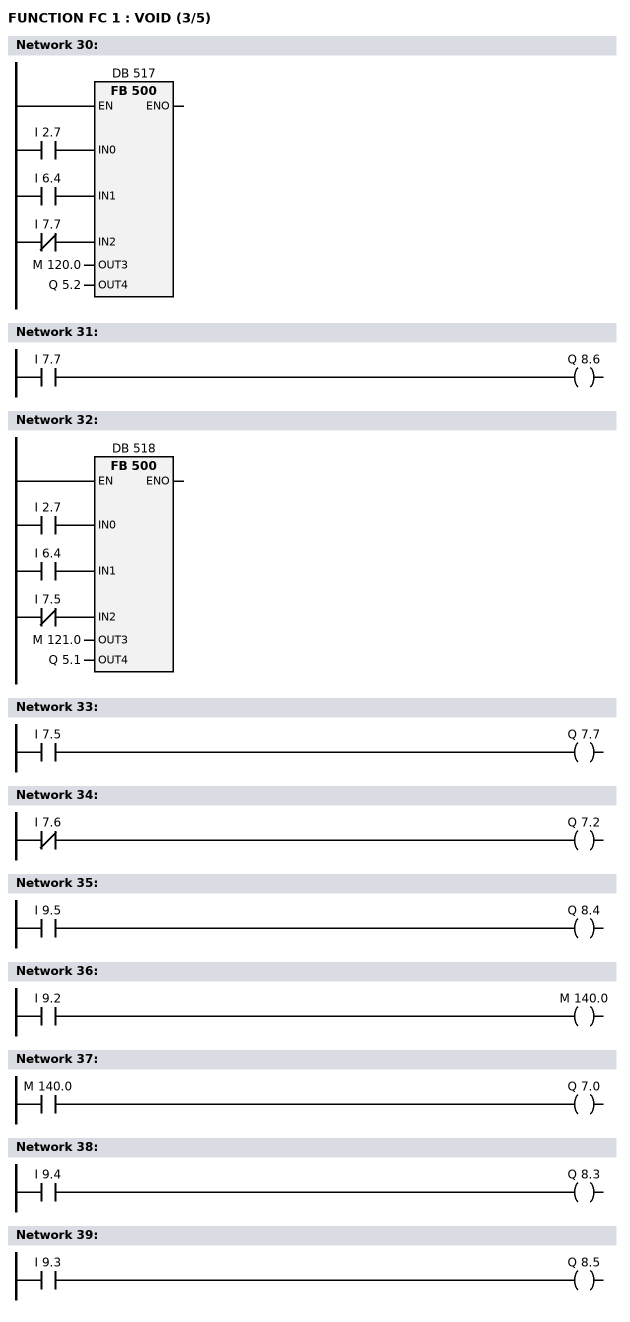

      A     I      2.7;
      =     L      0.0;
      BLD   103;
      A     I      6.4;
      =     L      0.1;
      BLD   103;
      AN    I      7.7;
      =     L      0.2;
      BLD   103;
      CALL FB   500 , DB   517 (
           IN0                      := L      0.0,
           IN1                      := L      0.1,
           IN2                      := L      0.2,
           OUT3                     := M    120.0,
           OUT4                     := Q      5.2);
      NOP   0;
NETWORK
TITLE =

      A     I      7.7;
      =     Q      8.6;
NETWORK
TITLE =

      A     I      2.7;
      =     L      0.0;
      BLD   103;
      A     I      6.4;
      =     L      0.1;
      BLD   103;
      AN    I      7.5;
      =     L      0.2;
      BLD   103;
      CALL FB   500 , DB   518 (
           IN0                      := L      0.0,
           IN1                      := L      0.1,
           IN2                      := L      0.2,
           OUT3                     := M    121.0,
           OUT4                     := Q      5.1);
      NOP   0;
NETWORK
TITLE =

      A     I      7.5;
      =     Q      7.7;
NETWORK
TITLE =

      AN    I      7.6;
      =     Q      7.2;
NETWORK
TITLE =

      A     I      9.5;
      =     Q      8.4;
NETWORK
TITLE =

      A     I      9.2;
      =     M    140.0;
NETWORK
TITLE =

      A     M    140.0;
      =     Q      7.0;
NETWORK
TITLE =

      A     I      9.4;
      =     Q      8.3;
NETWORK
TITLE =

      A     I      9.3;
      =     Q      8.5;
NETWORK
TITLE =
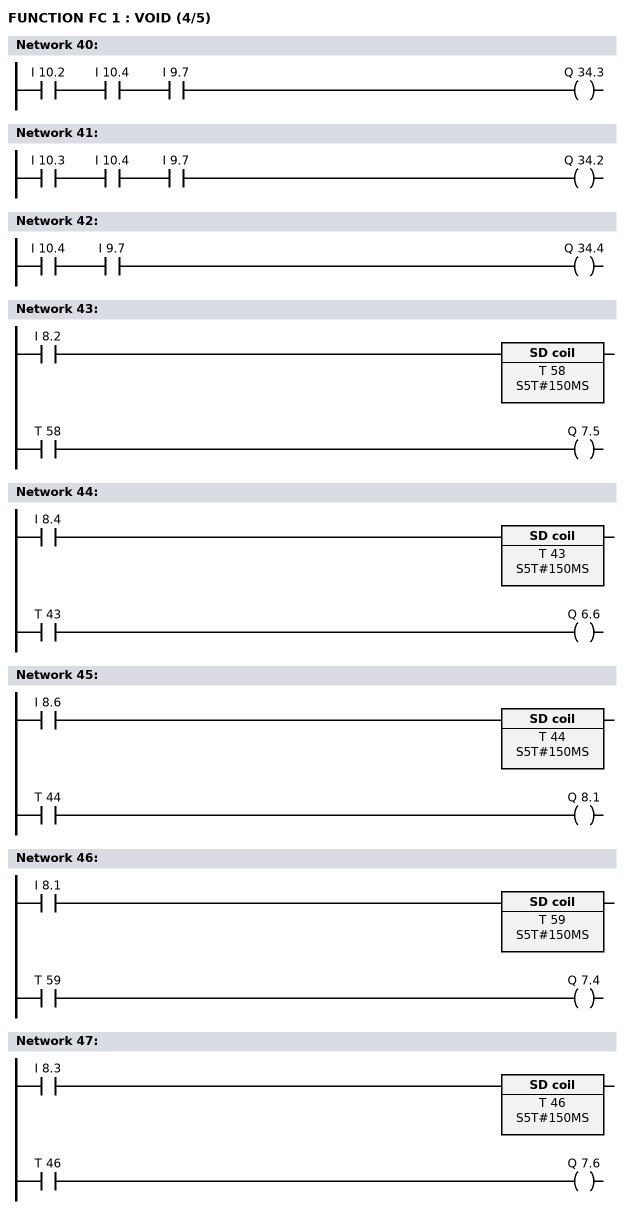

      A     I     10.2;
      A     I     10.4;
      A     I      9.7;
      =     Q     34.3;
NETWORK
TITLE =

      A     I     10.3;
      A     I     10.4;
      A     I      9.7;
      =     Q     34.2;
NETWORK
TITLE =

      A     I     10.4;
      A     I      9.7;
      =     Q     34.4;
NETWORK
TITLE =

      A     I      8.2;
      L     S5T#150MS;
      SD    T     58;
      NOP   0;
      NOP   0;
      NOP   0;
      A     T     58;
      =     Q      7.5;
NETWORK
TITLE =

      A     I      8.4;
      L     S5T#150MS;
      SD    T     43;
      NOP   0;
      NOP   0;
      NOP   0;
      A     T     43;
      =     Q      6.6;
NETWORK
TITLE =

      A     I      8.6;
      L     S5T#150MS;
      SD    T     44;
      NOP   0;
      NOP   0;
      NOP   0;
      A     T     44;
      =     Q      8.1;
NETWORK
TITLE =

      A     I      8.1;
      L     S5T#150MS;
      SD    T     59;
      NOP   0;
      NOP   0;
      NOP   0;
      A     T     59;
      =     Q      7.4;
NETWORK
TITLE =

      A     I      8.3;
      L     S5T#150MS;
      SD    T     46;
      NOP   0;
      NOP   0;
      NOP   0;
      A     T     46;
      =     Q      7.6;
NETWORK
TITLE =
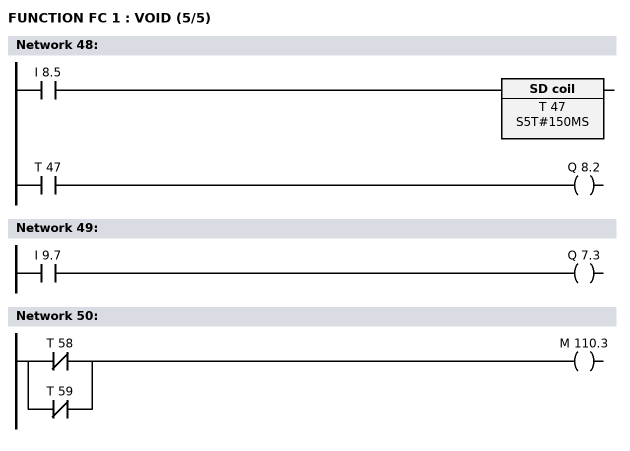

      A     I      8.5;
      L     S5T#150MS;
      SD    T     47;
      NOP   0;
      NOP   0;
      NOP   0;
      A     T     47;
      =     Q      8.2;
NETWORK
TITLE =

      A     I      9.7;
      =     Q      7.3;
NETWORK
TITLE =

      ON    T     58;
      ON    T     59;
      =     M    110.3;
END_FUNCTION

FUNCTION FC 2 : VOID
VERSION : 0.1

BEGIN
NETWORK
TITLE =
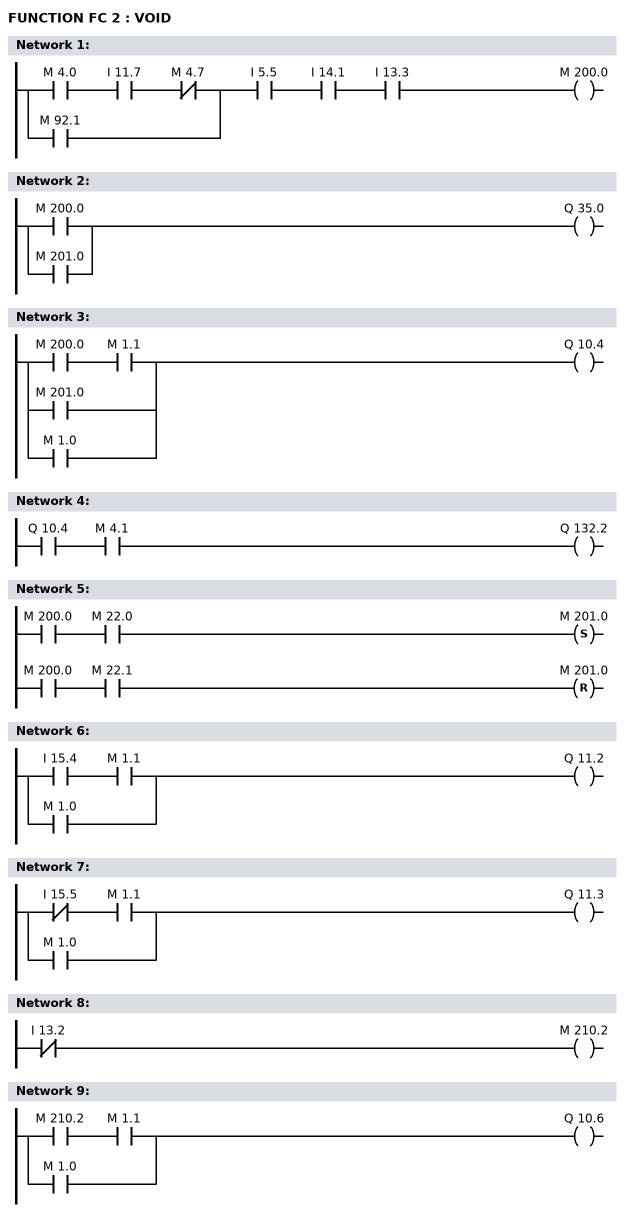

      A(    ;
      A     M      4.0;
      A     I     11.7;
      AN    M      4.7;
      O     M     92.1;
      )     ;
      A     I      5.5;
      A     I     14.1;
      A     I     13.3;
      =     M    200.0;
NETWORK
TITLE =

      O     M    200.0;
      O     M    201.0;
      =     Q     35.0;
NETWORK
TITLE =

      A     M    200.0;
      A     M      1.1;
      O     M    201.0;
      O     M      1.0;
      =     Q     10.4;
NETWORK
TITLE =

      A     Q     10.4;
      A     M      4.1;
      =     Q    132.2;
NETWORK
TITLE =

      A     M    200.0;
      A     M     22.0;
      S     M    201.0;
      A     M    200.0;
      A     M     22.1;
      R     M    201.0;
      NOP   0;
NETWORK
TITLE =

      A     I     15.4;
      A     M      1.1;
      O     M      1.0;
      =     Q     11.2;
NETWORK
TITLE =

      AN    I     15.5;
      A     M      1.1;
      O     M      1.0;
      =     Q     11.3;
NETWORK
TITLE =

      AN    I     13.2;
      =     M    210.2;
NETWORK
TITLE =

      A     M    210.2;
      A     M      1.1;
      O     M      1.0;
      =     Q     10.6;
NETWORK
TITLE =

      O(    ;
      A     I     12.3;
      L     S5T#150MS;
      SD    T     70;
      NOP   0;
      NOP   0;
      NOP   0;
      A     T     70;
      )     ;
      O     M      1.0;
      =     Q     10.3;
NETWORK
TITLE =
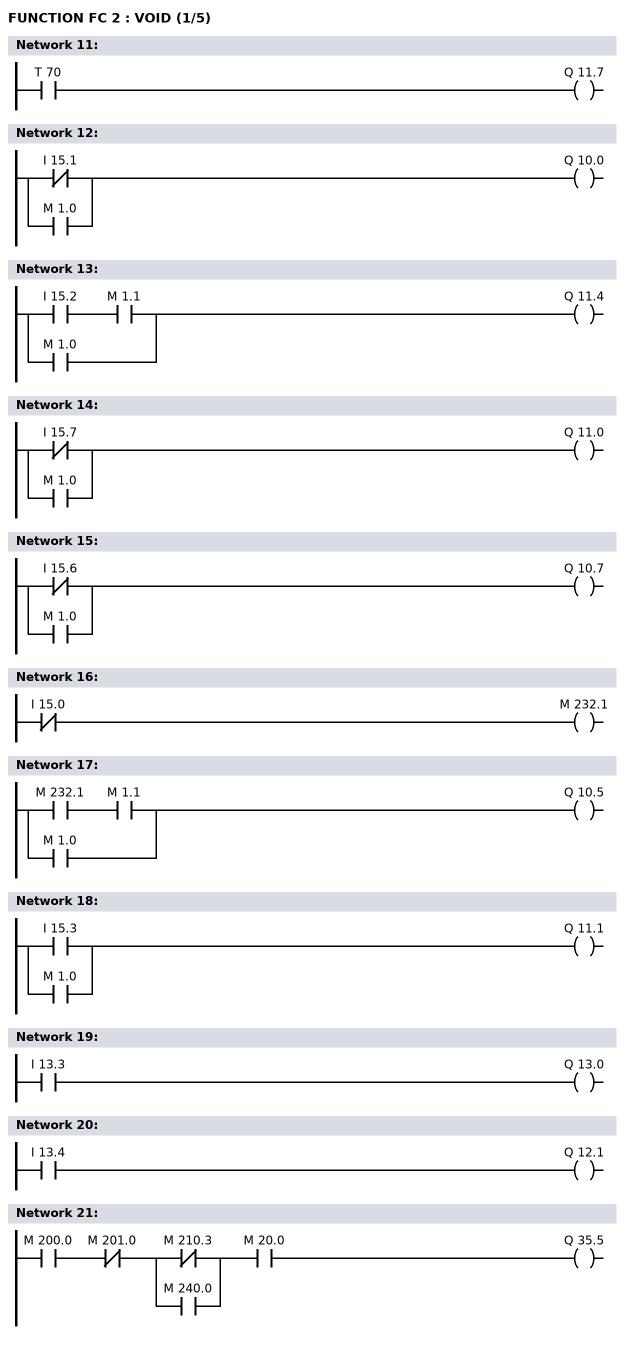

      A     T     70;
      =     Q     11.7;
NETWORK
TITLE =

      ON    I     15.1;
      O     M      1.0;
      =     Q     10.0;
NETWORK
TITLE =

      A     I     15.2;
      A     M      1.1;
      O     M      1.0;
      =     Q     11.4;
NETWORK
TITLE =

      ON    I     15.7;
      O     M      1.0;
      =     Q     11.0;
NETWORK
TITLE =

      ON    I     15.6;
      O     M      1.0;
      =     Q     10.7;
NETWORK
TITLE =

      AN    I     15.0;
      =     M    232.1;
NETWORK
TITLE =

      A     M    232.1;
      A     M      1.1;
      O     M      1.0;
      =     Q     10.5;
NETWORK
TITLE =

      O     I     15.3;
      O     M      1.0;
      =     Q     11.1;
NETWORK
TITLE =

      A     I     13.3;
      =     Q     13.0;
NETWORK
TITLE =

      A     I     13.4;
      =     Q     12.1;
NETWORK
TITLE =

      A     M    200.0;
      AN    M    201.0;
      A(    ;
      ON    M    210.3;
      O     M    240.0;
      )     ;
      A     M     20.0;
      =     Q     35.5;
NETWORK
TITLE =
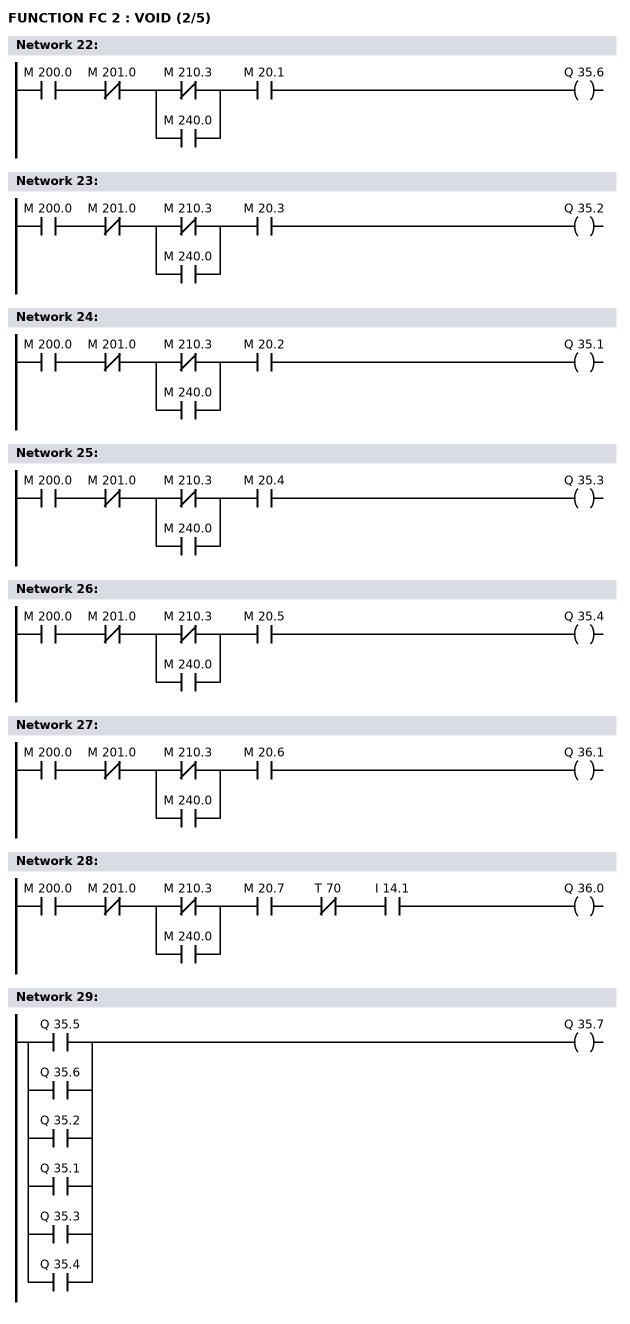

      A     M    200.0;
      AN    M    201.0;
      A(    ;
      ON    M    210.3;
      O     M    240.0;
      )     ;
      A     M     20.1;
      =     Q     35.6;
NETWORK
TITLE =

      A     M    200.0;
      AN    M    201.0;
      A(    ;
      ON    M    210.3;
      O     M    240.0;
      )     ;
      A     M     20.3;
      =     Q     35.2;
NETWORK
TITLE =

      A     M    200.0;
      AN    M    201.0;
      A(    ;
      ON    M    210.3;
      O     M    240.0;
      )     ;
      A     M     20.2;
      =     Q     35.1;
NETWORK
TITLE =

      A     M    200.0;
      AN    M    201.0;
      A(    ;
      ON    M    210.3;
      O     M    240.0;
      )     ;
      A     M     20.4;
      =     Q     35.3;
NETWORK
TITLE =

      A     M    200.0;
      AN    M    201.0;
      A(    ;
      ON    M    210.3;
      O     M    240.0;
      )     ;
      A     M     20.5;
      =     Q     35.4;
NETWORK
TITLE =

      A     M    200.0;
      AN    M    201.0;
      A(    ;
      ON    M    210.3;
      O     M    240.0;
      )     ;
      A     M     20.6;
      =     Q     36.1;
NETWORK
TITLE =

      A     M    200.0;
      AN    M    201.0;
      A(    ;
      ON    M    210.3;
      O     M    240.0;
      )     ;
      A     M     20.7;
      AN    T     70;
      A     I     14.1;
      =     Q     36.0;
NETWORK
TITLE =

      O     Q     35.5;
      O     Q     35.6;
      O     Q     35.2;
      O     Q     35.1;
      O     Q     35.3;
      O     Q     35.4;
      =     Q     35.7;
NETWORK
TITLE =
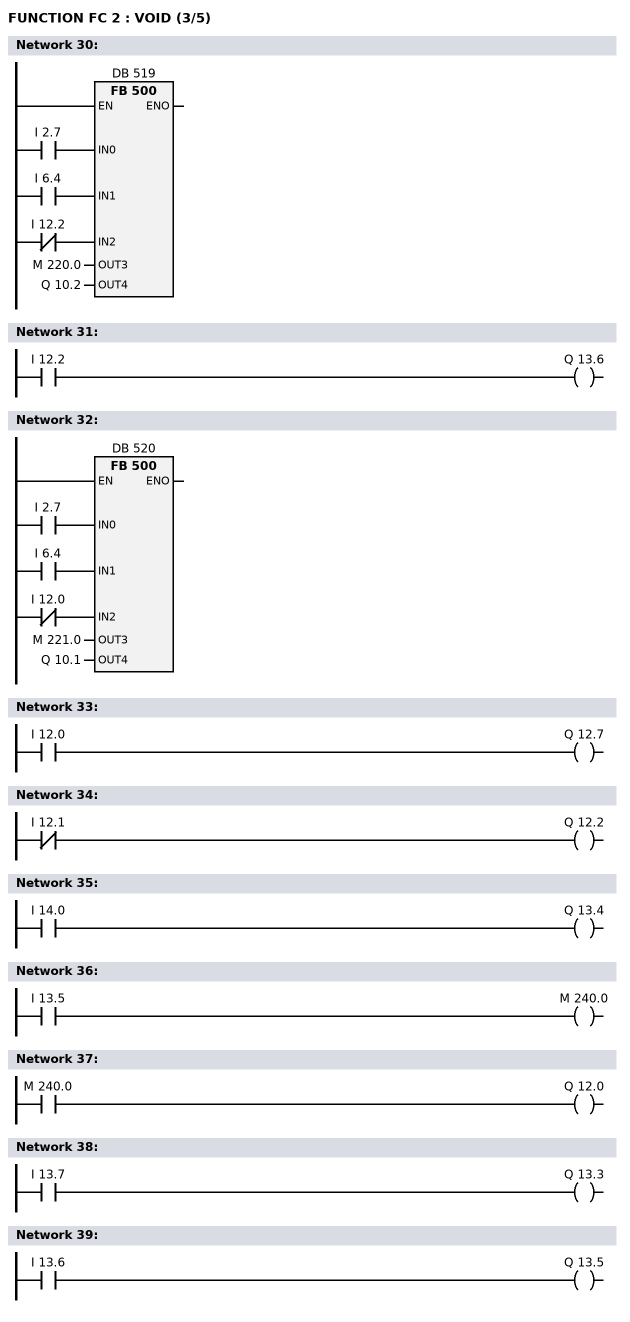

      A     I      2.7;
      =     L      0.0;
      BLD   103;
      A     I      6.4;
      =     L      0.1;
      BLD   103;
      AN    I     12.2;
      =     L      0.2;
      BLD   103;
      CALL FB   500 , DB   519 (
           IN0                      := L      0.0,
           IN1                      := L      0.1,
           IN2                      := L      0.2,
           OUT3                     := M    220.0,
           OUT4                     := Q     10.2);
      NOP   0;
NETWORK
TITLE =

      A     I     12.2;
      =     Q     13.6;
NETWORK
TITLE =

      A     I      2.7;
      =     L      0.0;
      BLD   103;
      A     I      6.4;
      =     L      0.1;
      BLD   103;
      AN    I     12.0;
      =     L      0.2;
      BLD   103;
      CALL FB   500 , DB   520 (
           IN0                      := L      0.0,
           IN1                      := L      0.1,
           IN2                      := L      0.2,
           OUT3                     := M    221.0,
           OUT4                     := Q     10.1);
      NOP   0;
NETWORK
TITLE =

      A     I     12.0;
      =     Q     12.7;
NETWORK
TITLE =

      AN    I     12.1;
      =     Q     12.2;
NETWORK
TITLE =

      A     I     14.0;
      =     Q     13.4;
NETWORK
TITLE =

      A     I     13.5;
      =     M    240.0;
NETWORK
TITLE =

      A     M    240.0;
      =     Q     12.0;
NETWORK
TITLE =

      A     I     13.7;
      =     Q     13.3;
NETWORK
TITLE =

      A     I     13.6;
      =     Q     13.5;
NETWORK
TITLE =
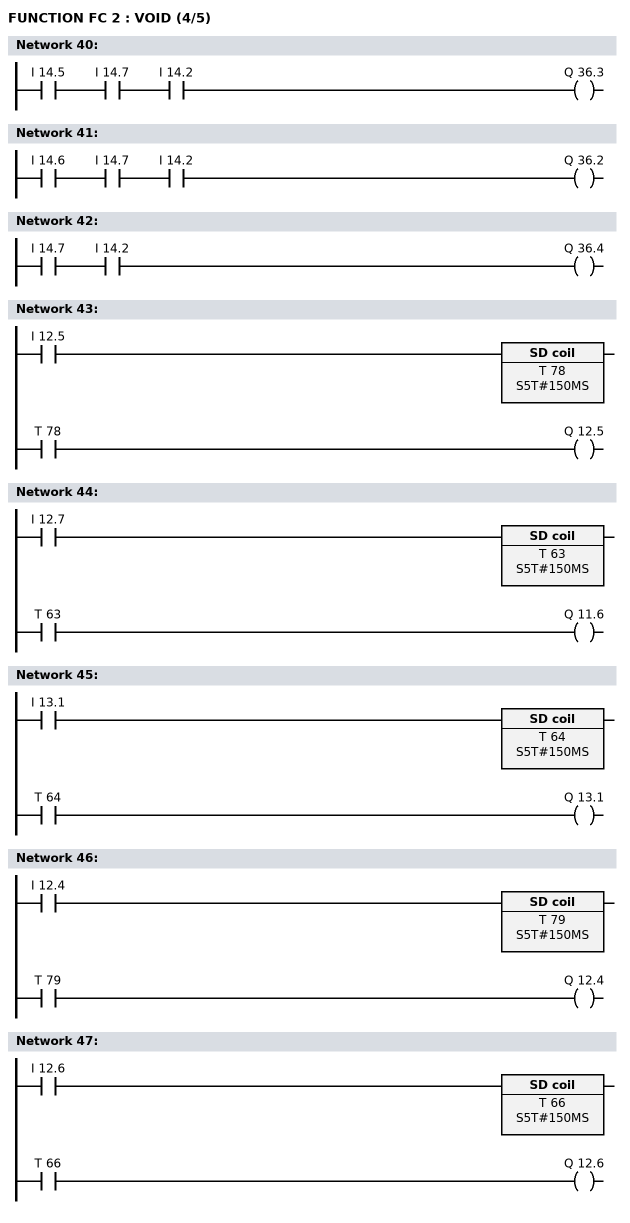

      A     I     14.5;
      A     I     14.7;
      A     I     14.2;
      =     Q     36.3;
NETWORK
TITLE =

      A     I     14.6;
      A     I     14.7;
      A     I     14.2;
      =     Q     36.2;
NETWORK
TITLE =

      A     I     14.7;
      A     I     14.2;
      =     Q     36.4;
NETWORK
TITLE =

      A     I     12.5;
      L     S5T#150MS;
      SD    T     78;
      NOP   0;
      NOP   0;
      NOP   0;
      A     T     78;
      =     Q     12.5;
NETWORK
TITLE =

      A     I     12.7;
      L     S5T#150MS;
      SD    T     63;
      NOP   0;
      NOP   0;
      NOP   0;
      A     T     63;
      =     Q     11.6;
NETWORK
TITLE =

      A     I     13.1;
      L     S5T#150MS;
      SD    T     64;
      NOP   0;
      NOP   0;
      NOP   0;
      A     T     64;
      =     Q     13.1;
NETWORK
TITLE =

      A     I     12.4;
      L     S5T#150MS;
      SD    T     79;
      NOP   0;
      NOP   0;
      NOP   0;
      A     T     79;
      =     Q     12.4;
NETWORK
TITLE =

      A     I     12.6;
      L     S5T#150MS;
      SD    T     66;
      NOP   0;
      NOP   0;
      NOP   0;
      A     T     66;
      =     Q     12.6;
NETWORK
TITLE =
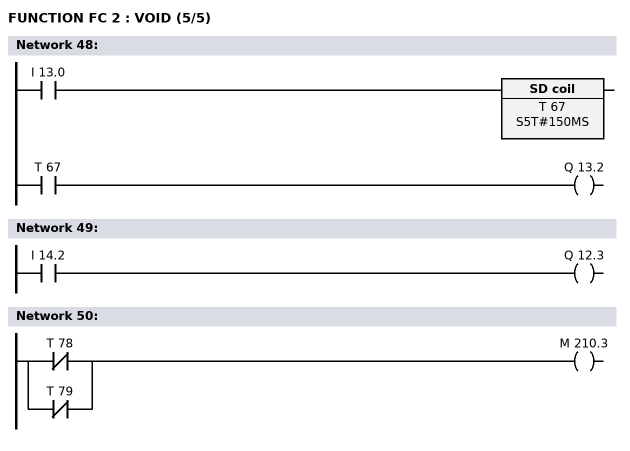

      A     I     13.0;
      L     S5T#150MS;
      SD    T     67;
      NOP   0;
      NOP   0;
      NOP   0;
      A     T     67;
      =     Q     13.2;
NETWORK
TITLE =

      A     I     14.2;
      =     Q     12.3;
NETWORK
TITLE =

      ON    T     78;
      ON    T     79;
      =     M    210.3;
END_FUNCTION

FUNCTION FC 3 : VOID
VERSION : 0.1

BEGIN
NETWORK
TITLE =
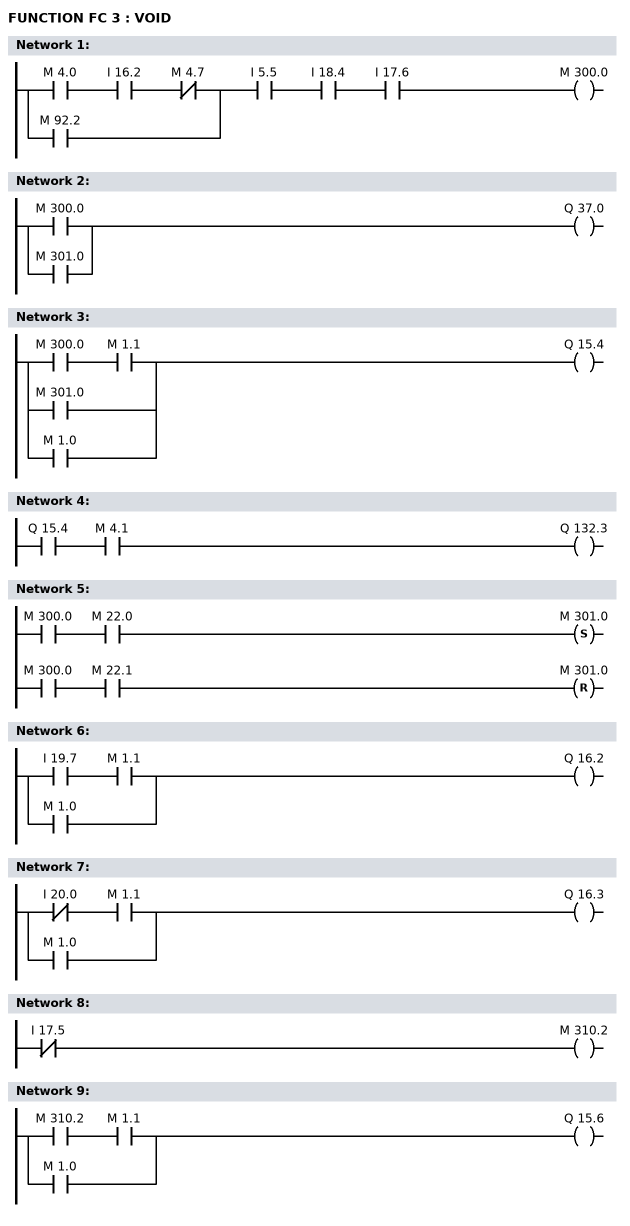

      A(    ;
      A     M      4.0;
      A     I     16.2;
      AN    M      4.7;
      O     M     92.2;
      )     ;
      A     I      5.5;
      A     I     18.4;
      A     I     17.6;
      =     M    300.0;
NETWORK
TITLE =

      O     M    300.0;
      O     M    301.0;
      =     Q     37.0;
NETWORK
TITLE =

      A     M    300.0;
      A     M      1.1;
      O     M    301.0;
      O     M      1.0;
      =     Q     15.4;
NETWORK
TITLE =

      A     Q     15.4;
      A     M      4.1;
      =     Q    132.3;
NETWORK
TITLE =

      A     M    300.0;
      A     M     22.0;
      S     M    301.0;
      A     M    300.0;
      A     M     22.1;
      R     M    301.0;
      NOP   0;
NETWORK
TITLE =

      A     I     19.7;
      A     M      1.1;
      O     M      1.0;
      =     Q     16.2;
NETWORK
TITLE =

      AN    I     20.0;
      A     M      1.1;
      O     M      1.0;
      =     Q     16.3;
NETWORK
TITLE =

      AN    I     17.5;
      =     M    310.2;
NETWORK
TITLE =

      A     M    310.2;
      A     M      1.1;
      O     M      1.0;
      =     Q     15.6;
NETWORK
TITLE =

      O(    ;
      A     I     16.6;
      L     S5T#150MS;
      SD    T     90;
      NOP   0;
      NOP   0;
      NOP   0;
      A     T     90;
      )     ;
      O     M      1.0;
      =     Q     15.3;
NETWORK
TITLE =
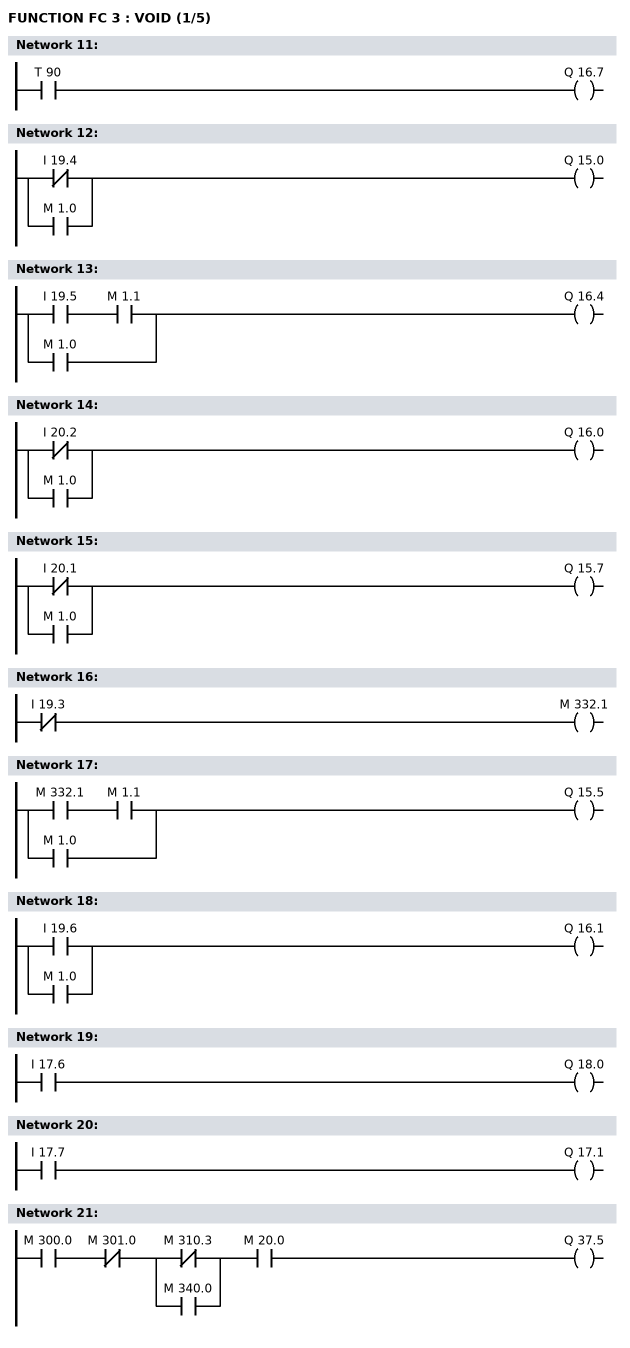

      A     T     90;
      =     Q     16.7;
NETWORK
TITLE =

      ON    I     19.4;
      O     M      1.0;
      =     Q     15.0;
NETWORK
TITLE =

      A     I     19.5;
      A     M      1.1;
      O     M      1.0;
      =     Q     16.4;
NETWORK
TITLE =

      ON    I     20.2;
      O     M      1.0;
      =     Q     16.0;
NETWORK
TITLE =

      ON    I     20.1;
      O     M      1.0;
      =     Q     15.7;
NETWORK
TITLE =

      AN    I     19.3;
      =     M    332.1;
NETWORK
TITLE =

      A     M    332.1;
      A     M      1.1;
      O     M      1.0;
      =     Q     15.5;
NETWORK
TITLE =

      O     I     19.6;
      O     M      1.0;
      =     Q     16.1;
NETWORK
TITLE =

      A     I     17.6;
      =     Q     18.0;
NETWORK
TITLE =

      A     I     17.7;
      =     Q     17.1;
NETWORK
TITLE =

      A     M    300.0;
      AN    M    301.0;
      A(    ;
      ON    M    310.3;
      O     M    340.0;
      )     ;
      A     M     20.0;
      =     Q     37.5;
NETWORK
TITLE =
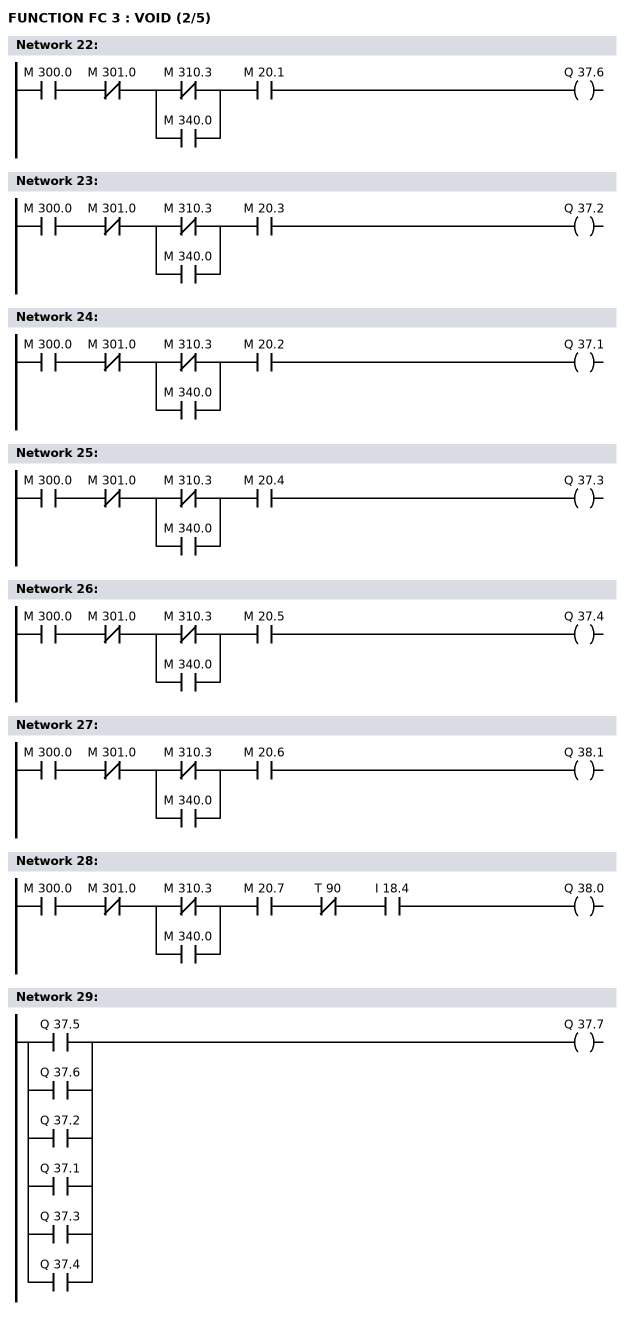

      A     M    300.0;
      AN    M    301.0;
      A(    ;
      ON    M    310.3;
      O     M    340.0;
      )     ;
      A     M     20.1;
      =     Q     37.6;
NETWORK
TITLE =

      A     M    300.0;
      AN    M    301.0;
      A(    ;
      ON    M    310.3;
      O     M    340.0;
      )     ;
      A     M     20.3;
      =     Q     37.2;
NETWORK
TITLE =

      A     M    300.0;
      AN    M    301.0;
      A(    ;
      ON    M    310.3;
      O     M    340.0;
      )     ;
      A     M     20.2;
      =     Q     37.1;
NETWORK
TITLE =

      A     M    300.0;
      AN    M    301.0;
      A(    ;
      ON    M    310.3;
      O     M    340.0;
      )     ;
      A     M     20.4;
      =     Q     37.3;
NETWORK
TITLE =

      A     M    300.0;
      AN    M    301.0;
      A(    ;
      ON    M    310.3;
      O     M    340.0;
      )     ;
      A     M     20.5;
      =     Q     37.4;
NETWORK
TITLE =

      A     M    300.0;
      AN    M    301.0;
      A(    ;
      ON    M    310.3;
      O     M    340.0;
      )     ;
      A     M     20.6;
      =     Q     38.1;
NETWORK
TITLE =

      A     M    300.0;
      AN    M    301.0;
      A(    ;
      ON    M    310.3;
      O     M    340.0;
      )     ;
      A     M     20.7;
      AN    T     90;
      A     I     18.4;
      =     Q     38.0;
NETWORK
TITLE =

      O     Q     37.5;
      O     Q     37.6;
      O     Q     37.2;
      O     Q     37.1;
      O     Q     37.3;
      O     Q     37.4;
      =     Q     37.7;
NETWORK
TITLE =
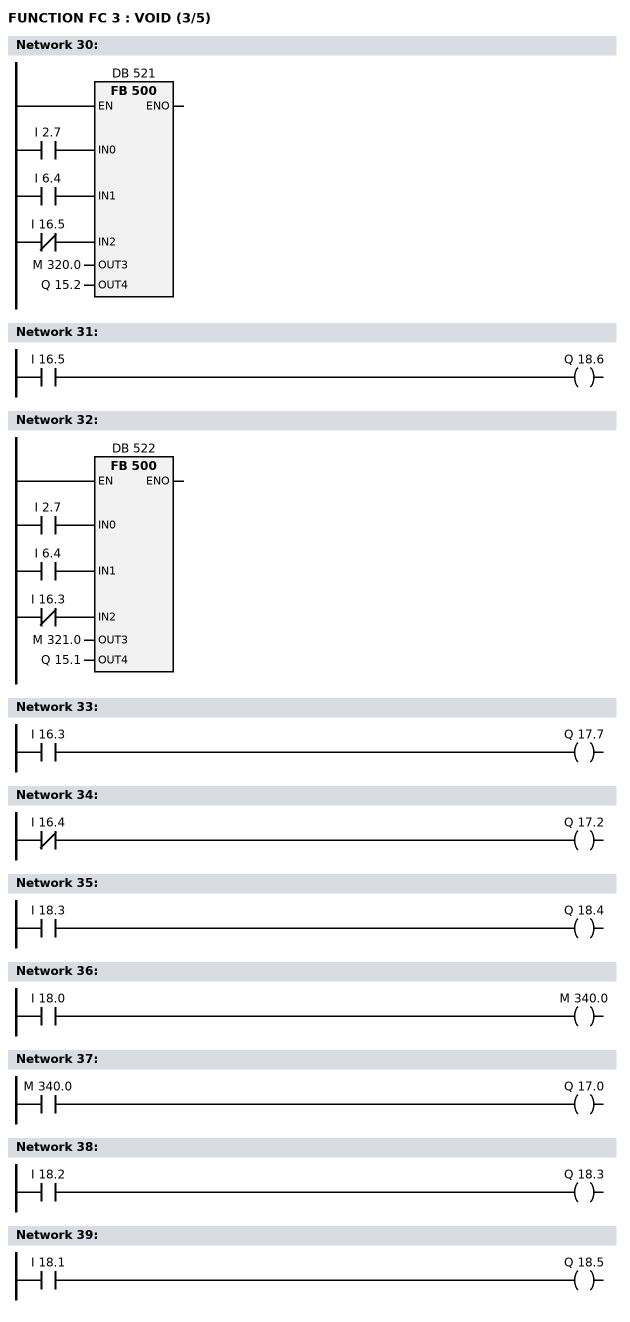

      A     I      2.7;
      =     L      0.0;
      BLD   103;
      A     I      6.4;
      =     L      0.1;
      BLD   103;
      AN    I     16.5;
      =     L      0.2;
      BLD   103;
      CALL FB   500 , DB   521 (
           IN0                      := L      0.0,
           IN1                      := L      0.1,
           IN2                      := L      0.2,
           OUT3                     := M    320.0,
           OUT4                     := Q     15.2);
      NOP   0;
NETWORK
TITLE =

      A     I     16.5;
      =     Q     18.6;
NETWORK
TITLE =

      A     I      2.7;
      =     L      0.0;
      BLD   103;
      A     I      6.4;
      =     L      0.1;
      BLD   103;
      AN    I     16.3;
      =     L      0.2;
      BLD   103;
      CALL FB   500 , DB   522 (
           IN0                      := L      0.0,
           IN1                      := L      0.1,
           IN2                      := L      0.2,
           OUT3                     := M    321.0,
           OUT4                     := Q     15.1);
      NOP   0;
NETWORK
TITLE =

      A     I     16.3;
      =     Q     17.7;
NETWORK
TITLE =

      AN    I     16.4;
      =     Q     17.2;
NETWORK
TITLE =

      A     I     18.3;
      =     Q     18.4;
NETWORK
TITLE =

      A     I     18.0;
      =     M    340.0;
NETWORK
TITLE =

      A     M    340.0;
      =     Q     17.0;
NETWORK
TITLE =

      A     I     18.2;
      =     Q     18.3;
NETWORK
TITLE =

      A     I     18.1;
      =     Q     18.5;
NETWORK
TITLE =
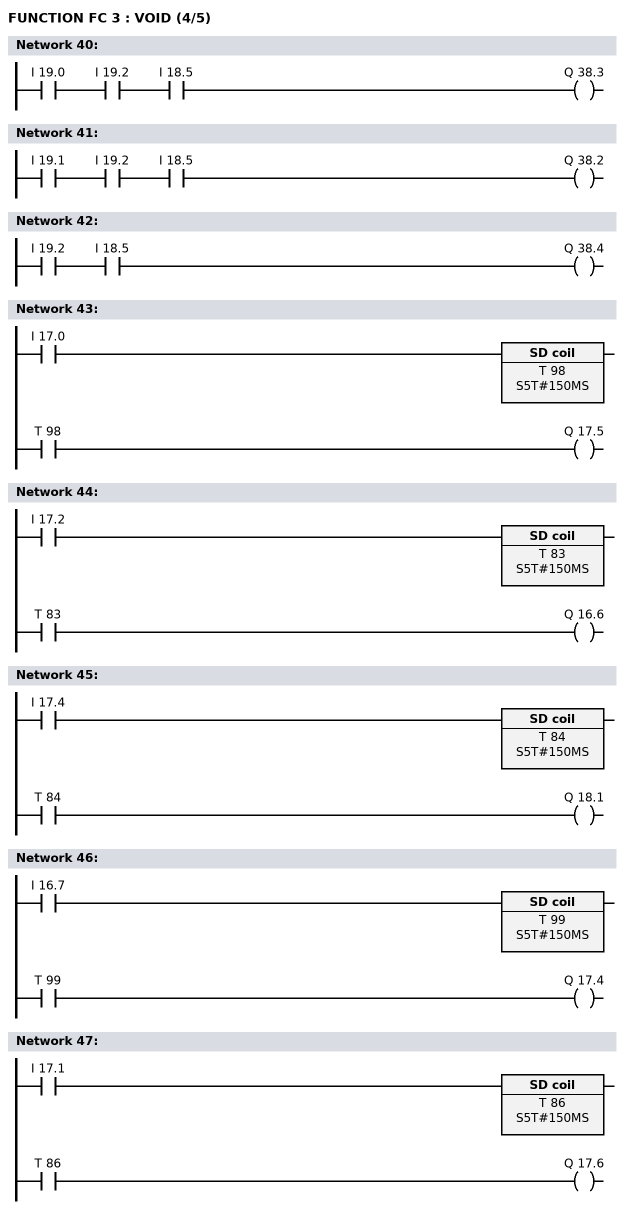

      A     I     19.0;
      A     I     19.2;
      A     I     18.5;
      =     Q     38.3;
NETWORK
TITLE =

      A     I     19.1;
      A     I     19.2;
      A     I     18.5;
      =     Q     38.2;
NETWORK
TITLE =

      A     I     19.2;
      A     I     18.5;
      =     Q     38.4;
NETWORK
TITLE =

      A     I     17.0;
      L     S5T#150MS;
      SD    T     98;
      NOP   0;
      NOP   0;
      NOP   0;
      A     T     98;
      =     Q     17.5;
NETWORK
TITLE =

      A     I     17.2;
      L     S5T#150MS;
      SD    T     83;
      NOP   0;
      NOP   0;
      NOP   0;
      A     T     83;
      =     Q     16.6;
NETWORK
TITLE =

      A     I     17.4;
      L     S5T#150MS;
      SD    T     84;
      NOP   0;
      NOP   0;
      NOP   0;
      A     T     84;
      =     Q     18.1;
NETWORK
TITLE =

      A     I     16.7;
      L     S5T#150MS;
      SD    T     99;
      NOP   0;
      NOP   0;
      NOP   0;
      A     T     99;
      =     Q     17.4;
NETWORK
TITLE =

      A     I     17.1;
      L     S5T#150MS;
      SD    T     86;
      NOP   0;
      NOP   0;
      NOP   0;
      A     T     86;
      =     Q     17.6;
NETWORK
TITLE =
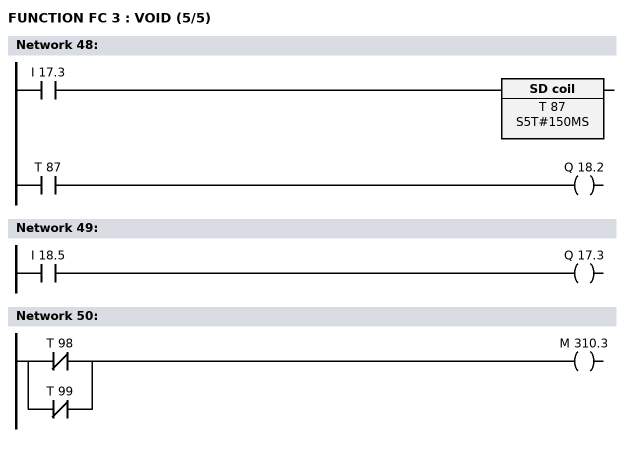

      A     I     17.3;
      L     S5T#150MS;
      SD    T     87;
      NOP   0;
      NOP   0;
      NOP   0;
      A     T     87;
      =     Q     18.2;
NETWORK
TITLE =

      A     I     18.5;
      =     Q     17.3;
NETWORK
TITLE =

      ON    T     98;
      ON    T     99;
      =     M    310.3;
END_FUNCTION

FUNCTION FC 4 : VOID
VERSION : 0.1

BEGIN
NETWORK
TITLE =
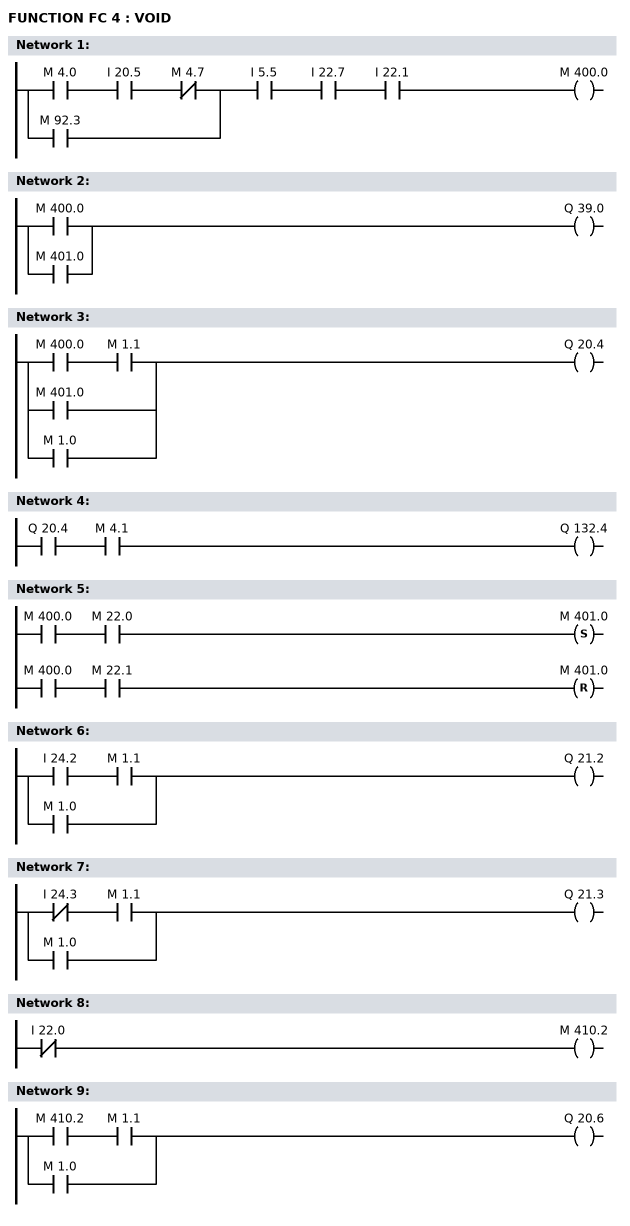

      A(    ;
      A     M      4.0;
      A     I     20.5;
      AN    M      4.7;
      O     M     92.3;
      )     ;
      A     I      5.5;
      A     I     22.7;
      A     I     22.1;
      =     M    400.0;
NETWORK
TITLE =

      O     M    400.0;
      O     M    401.0;
      =     Q     39.0;
NETWORK
TITLE =

      A     M    400.0;
      A     M      1.1;
      O     M    401.0;
      O     M      1.0;
      =     Q     20.4;
NETWORK
TITLE =

      A     Q     20.4;
      A     M      4.1;
      =     Q    132.4;
NETWORK
TITLE =

      A     M    400.0;
      A     M     22.0;
      S     M    401.0;
      A     M    400.0;
      A     M     22.1;
      R     M    401.0;
      NOP   0;
NETWORK
TITLE =

      A     I     24.2;
      A     M      1.1;
      O     M      1.0;
      =     Q     21.2;
NETWORK
TITLE =

      AN    I     24.3;
      A     M      1.1;
      O     M      1.0;
      =     Q     21.3;
NETWORK
TITLE =

      AN    I     22.0;
      =     M    410.2;
NETWORK
TITLE =

      A     M    410.2;
      A     M      1.1;
      O     M      1.0;
      =     Q     20.6;
NETWORK
TITLE =

      O(    ;
      A     I     21.1;
      L     S5T#150MS;
      SD    T    110;
      NOP   0;
      NOP   0;
      NOP   0;
      A     T    110;
      )     ;
      O     M      1.0;
      =     Q     20.3;
NETWORK
TITLE =
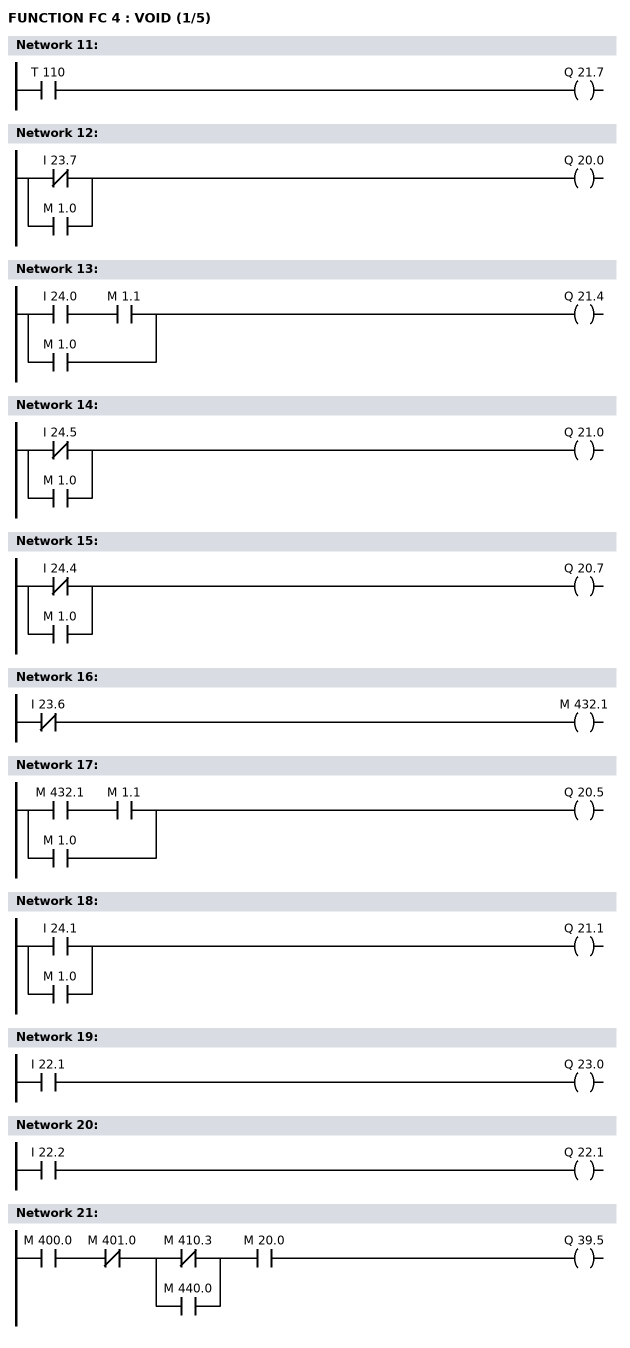

      A     T    110;
      =     Q     21.7;
NETWORK
TITLE =

      ON    I     23.7;
      O     M      1.0;
      =     Q     20.0;
NETWORK
TITLE =

      A     I     24.0;
      A     M      1.1;
      O     M      1.0;
      =     Q     21.4;
NETWORK
TITLE =

      ON    I     24.5;
      O     M      1.0;
      =     Q     21.0;
NETWORK
TITLE =

      ON    I     24.4;
      O     M      1.0;
      =     Q     20.7;
NETWORK
TITLE =

      AN    I     23.6;
      =     M    432.1;
NETWORK
TITLE =

      A     M    432.1;
      A     M      1.1;
      O     M      1.0;
      =     Q     20.5;
NETWORK
TITLE =

      O     I     24.1;
      O     M      1.0;
      =     Q     21.1;
NETWORK
TITLE =

      A     I     22.1;
      =     Q     23.0;
NETWORK
TITLE =

      A     I     22.2;
      =     Q     22.1;
NETWORK
TITLE =

      A     M    400.0;
      AN    M    401.0;
      A(    ;
      ON    M    410.3;
      O     M    440.0;
      )     ;
      A     M     20.0;
      =     Q     39.5;
NETWORK
TITLE =
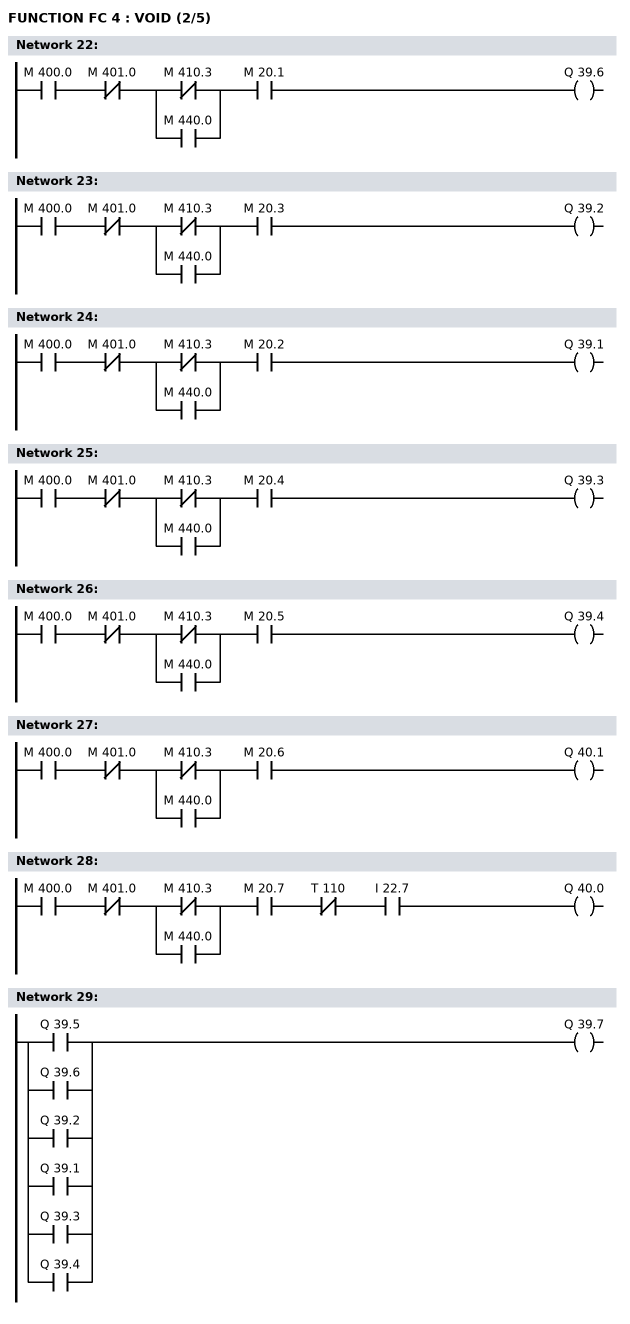

      A     M    400.0;
      AN    M    401.0;
      A(    ;
      ON    M    410.3;
      O     M    440.0;
      )     ;
      A     M     20.1;
      =     Q     39.6;
NETWORK
TITLE =

      A     M    400.0;
      AN    M    401.0;
      A(    ;
      ON    M    410.3;
      O     M    440.0;
      )     ;
      A     M     20.3;
      =     Q     39.2;
NETWORK
TITLE =

      A     M    400.0;
      AN    M    401.0;
      A(    ;
      ON    M    410.3;
      O     M    440.0;
      )     ;
      A     M     20.2;
      =     Q     39.1;
NETWORK
TITLE =

      A     M    400.0;
      AN    M    401.0;
      A(    ;
      ON    M    410.3;
      O     M    440.0;
      )     ;
      A     M     20.4;
      =     Q     39.3;
NETWORK
TITLE =

      A     M    400.0;
      AN    M    401.0;
      A(    ;
      ON    M    410.3;
      O     M    440.0;
      )     ;
      A     M     20.5;
      =     Q     39.4;
NETWORK
TITLE =

      A     M    400.0;
      AN    M    401.0;
      A(    ;
      ON    M    410.3;
      O     M    440.0;
      )     ;
      A     M     20.6;
      =     Q     40.1;
NETWORK
TITLE =

      A     M    400.0;
      AN    M    401.0;
      A(    ;
      ON    M    410.3;
      O     M    440.0;
      )     ;
      A     M     20.7;
      AN    T    110;
      A     I     22.7;
      =     Q     40.0;
NETWORK
TITLE =

      O     Q     39.5;
      O     Q     39.6;
      O     Q     39.2;
      O     Q     39.1;
      O     Q     39.3;
      O     Q     39.4;
      =     Q     39.7;
NETWORK
TITLE =
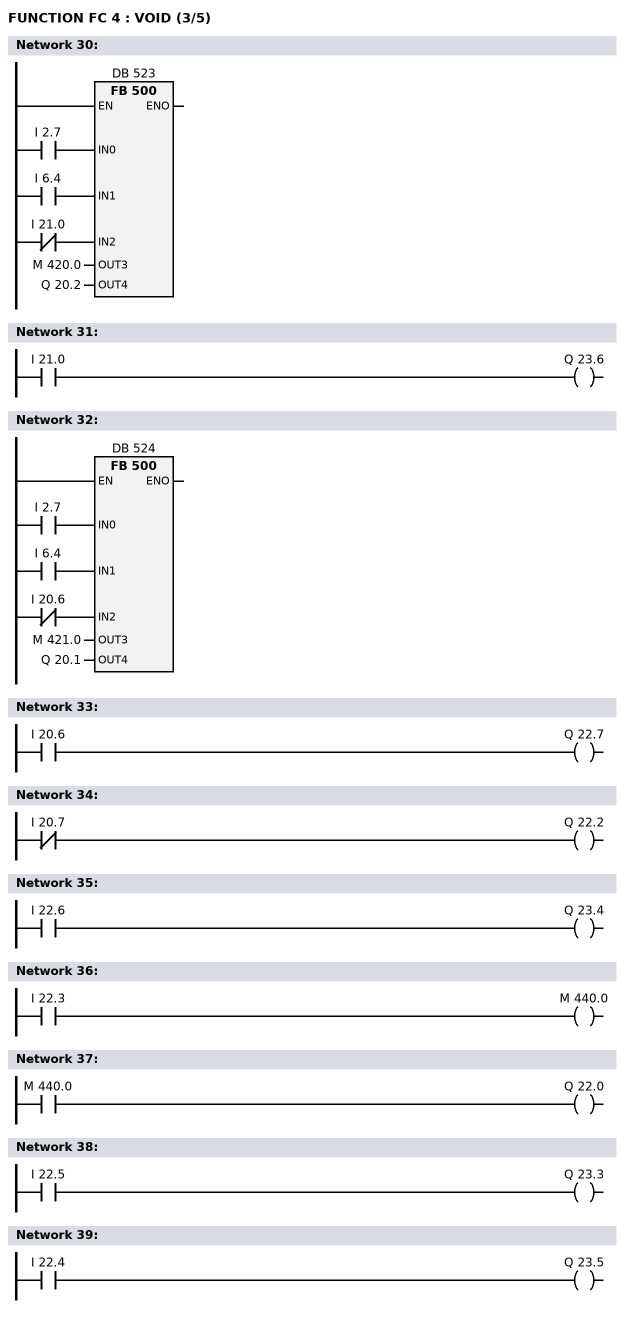

      A     I      2.7;
      =     L      0.0;
      BLD   103;
      A     I      6.4;
      =     L      0.1;
      BLD   103;
      AN    I     21.0;
      =     L      0.2;
      BLD   103;
      CALL FB   500 , DB   523 (
           IN0                      := L      0.0,
           IN1                      := L      0.1,
           IN2                      := L      0.2,
           OUT3                     := M    420.0,
           OUT4                     := Q     20.2);
      NOP   0;
NETWORK
TITLE =

      A     I     21.0;
      =     Q     23.6;
NETWORK
TITLE =

      A     I      2.7;
      =     L      0.0;
      BLD   103;
      A     I      6.4;
      =     L      0.1;
      BLD   103;
      AN    I     20.6;
      =     L      0.2;
      BLD   103;
      CALL FB   500 , DB   524 (
           IN0                      := L      0.0,
           IN1                      := L      0.1,
           IN2                      := L      0.2,
           OUT3                     := M    421.0,
           OUT4                     := Q     20.1);
      NOP   0;
NETWORK
TITLE =

      A     I     20.6;
      =     Q     22.7;
NETWORK
TITLE =

      AN    I     20.7;
      =     Q     22.2;
NETWORK
TITLE =

      A     I     22.6;
      =     Q     23.4;
NETWORK
TITLE =

      A     I     22.3;
      =     M    440.0;
NETWORK
TITLE =

      A     M    440.0;
      =     Q     22.0;
NETWORK
TITLE =

      A     I     22.5;
      =     Q     23.3;
NETWORK
TITLE =

      A     I     22.4;
      =     Q     23.5;
NETWORK
TITLE =
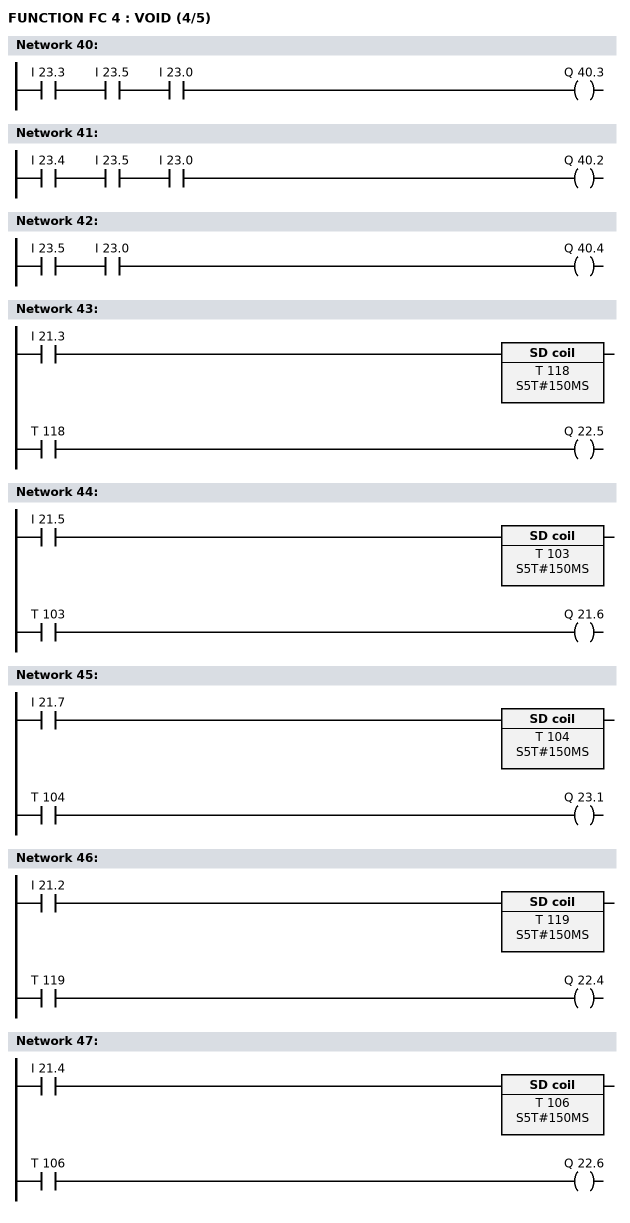

      A     I     23.3;
      A     I     23.5;
      A     I     23.0;
      =     Q     40.3;
NETWORK
TITLE =

      A     I     23.4;
      A     I     23.5;
      A     I     23.0;
      =     Q     40.2;
NETWORK
TITLE =

      A     I     23.5;
      A     I     23.0;
      =     Q     40.4;
NETWORK
TITLE =

      A     I     21.3;
      L     S5T#150MS;
      SD    T    118;
      NOP   0;
      NOP   0;
      NOP   0;
      A     T    118;
      =     Q     22.5;
NETWORK
TITLE =

      A     I     21.5;
      L     S5T#150MS;
      SD    T    103;
      NOP   0;
      NOP   0;
      NOP   0;
      A     T    103;
      =     Q     21.6;
NETWORK
TITLE =

      A     I     21.7;
      L     S5T#150MS;
      SD    T    104;
      NOP   0;
      NOP   0;
      NOP   0;
      A     T    104;
      =     Q     23.1;
NETWORK
TITLE =

      A     I     21.2;
      L     S5T#150MS;
      SD    T    119;
      NOP   0;
      NOP   0;
      NOP   0;
      A     T    119;
      =     Q     22.4;
NETWORK
TITLE =

      A     I     21.4;
      L     S5T#150MS;
      SD    T    106;
      NOP   0;
      NOP   0;
      NOP   0;
      A     T    106;
      =     Q     22.6;
NETWORK
TITLE =
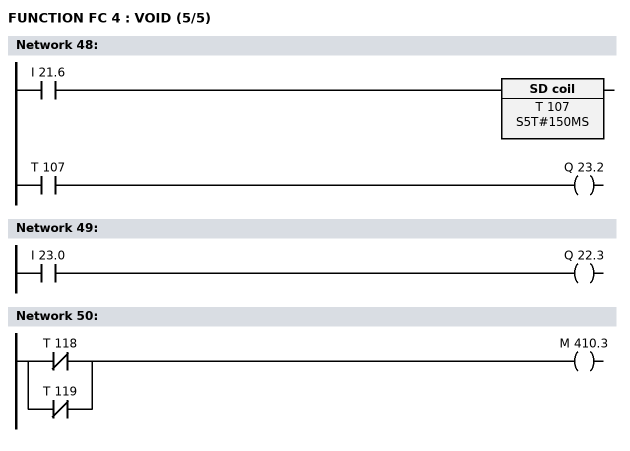

      A     I     21.6;
      L     S5T#150MS;
      SD    T    107;
      NOP   0;
      NOP   0;
      NOP   0;
      A     T    107;
      =     Q     23.2;
NETWORK
TITLE =

      A     I     23.0;
      =     Q     22.3;
NETWORK
TITLE =

      ON    T    118;
      ON    T    119;
      =     M    410.3;
END_FUNCTION

FUNCTION FC 11 : VOID
VERSION : 0.1

BEGIN
NETWORK
TITLE =
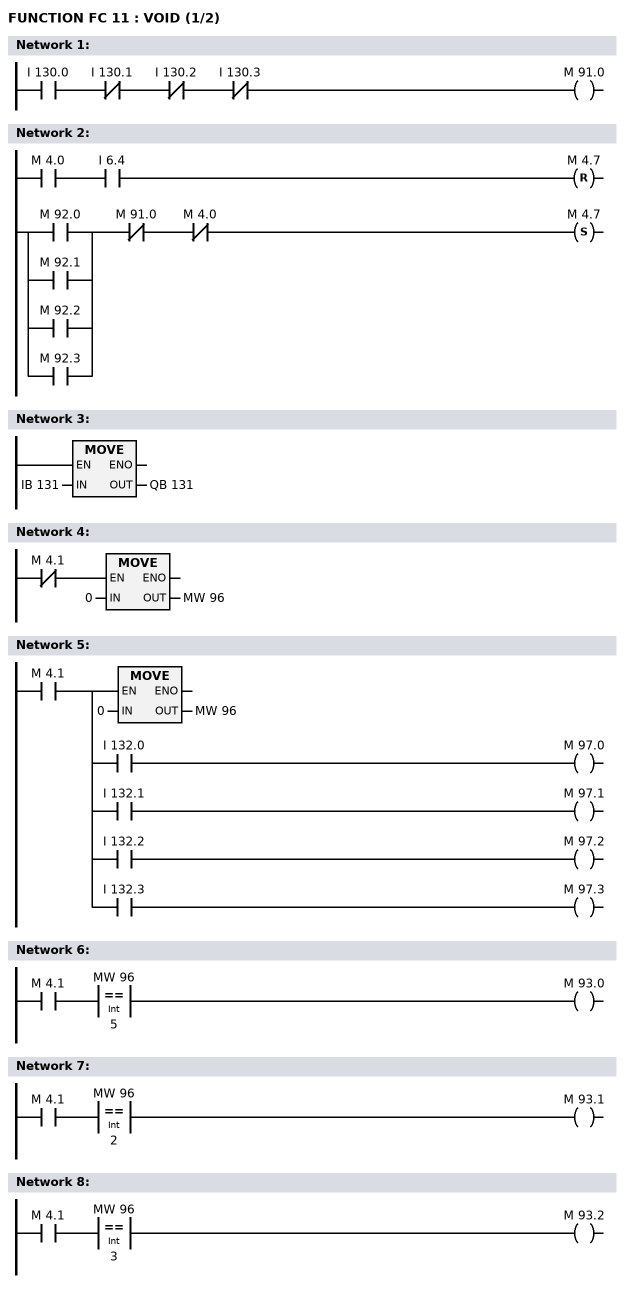

      A     I    130.0;
      AN    I    130.1;
      AN    I    130.2;
      AN    I    130.3;
      =     M     91.0;
NETWORK
TITLE =

      A     M      4.0;
      A     I      6.4;
      R     M      4.7;
      A(    ;
      O     M     92.0;
      O     M     92.1;
      O     M     92.2;
      O     M     92.3;
      )     ;
      AN    M     91.0;
      AN    M      4.0;
      S     M      4.7;
      NOP   0;
NETWORK
TITLE =

      L     IB   131;
      T     QB   131;
      NOP   0;
NETWORK
TITLE =

      AN    M      4.1;
      JNB   M001;
      L     0;
      T     MW    96;
M001: NOP   0;
NETWORK
TITLE =

      A     M      4.1;
      =     L      0.0;
      A     L      0.0;
      JNB   M002;
      L     0;
      T     MW    96;
M002: NOP   0;
      A     L      0.0;
      A     I    132.0;
      =     M     97.0;
      A     L      0.0;
      A     I    132.1;
      =     M     97.1;
      A     L      0.0;
      A     I    132.2;
      =     M     97.2;
      A     L      0.0;
      A     I    132.3;
      =     M     97.3;
NETWORK
TITLE =

      A     M      4.1;
      A(    ;
      L     MW    96;
      L     5;
      ==I   ;
      )     ;
      =     M     93.0;
NETWORK
TITLE =

      A     M      4.1;
      A(    ;
      L     MW    96;
      L     2;
      ==I   ;
      )     ;
      =     M     93.1;
NETWORK
TITLE =

      A     M      4.1;
      A(    ;
      L     MW    96;
      L     3;
      ==I   ;
      )     ;
      =     M     93.2;
NETWORK
TITLE =
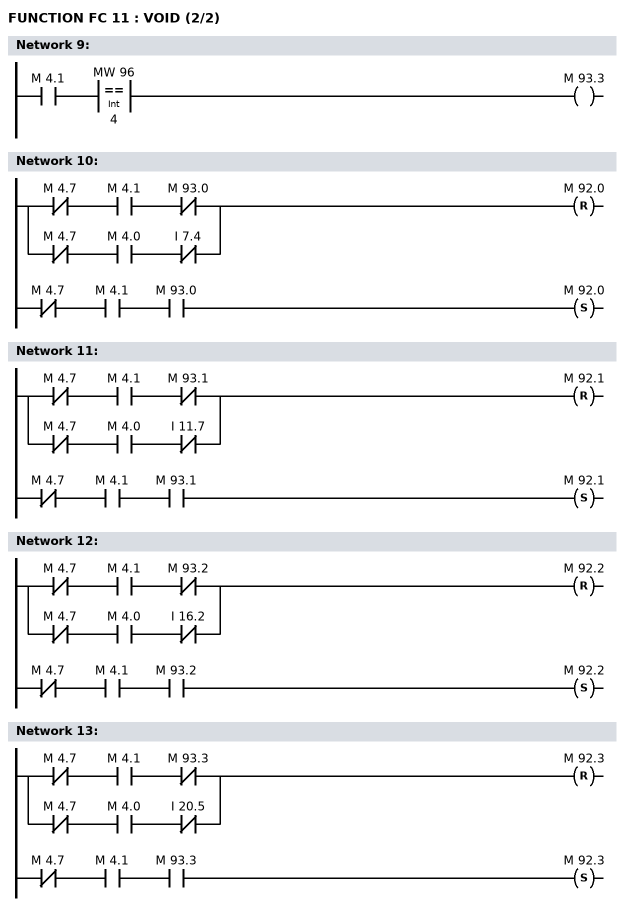

      A     M      4.1;
      A(    ;
      L     MW    96;
      L     4;
      ==I   ;
      )     ;
      =     M     93.3;
NETWORK
TITLE =

      A(    ;
      AN    M      4.7;
      A     M      4.1;
      AN    M     93.0;
      O     ;
      AN    M      4.7;
      A     M      4.0;
      AN    I      7.4;
      )     ;
      R     M     92.0;
      AN    M      4.7;
      A     M      4.1;
      A     M     93.0;
      S     M     92.0;
      NOP   0;
NETWORK
TITLE =

      A(    ;
      AN    M      4.7;
      A     M      4.1;
      AN    M     93.1;
      O     ;
      AN    M      4.7;
      A     M      4.0;
      AN    I     11.7;
      )     ;
      R     M     92.1;
      AN    M      4.7;
      A     M      4.1;
      A     M     93.1;
      S     M     92.1;
      NOP   0;
NETWORK
TITLE =

      A(    ;
      AN    M      4.7;
      A     M      4.1;
      AN    M     93.2;
      O     ;
      AN    M      4.7;
      A     M      4.0;
      AN    I     16.2;
      )     ;
      R     M     92.2;
      AN    M      4.7;
      A     M      4.1;
      A     M     93.2;
      S     M     92.2;
      NOP   0;
NETWORK
TITLE =

      A(    ;
      AN    M      4.7;
      A     M      4.1;
      AN    M     93.3;
      O     ;
      AN    M      4.7;
      A     M      4.0;
      AN    I     20.5;
      )     ;
      R     M     92.3;
      AN    M      4.7;
      A     M      4.1;
      A     M     93.3;
      S     M     92.3;
      NOP   0;
END_FUNCTION

FUNCTION FC 13 : VOID
VERSION : 0.1

BEGIN
NETWORK
TITLE =
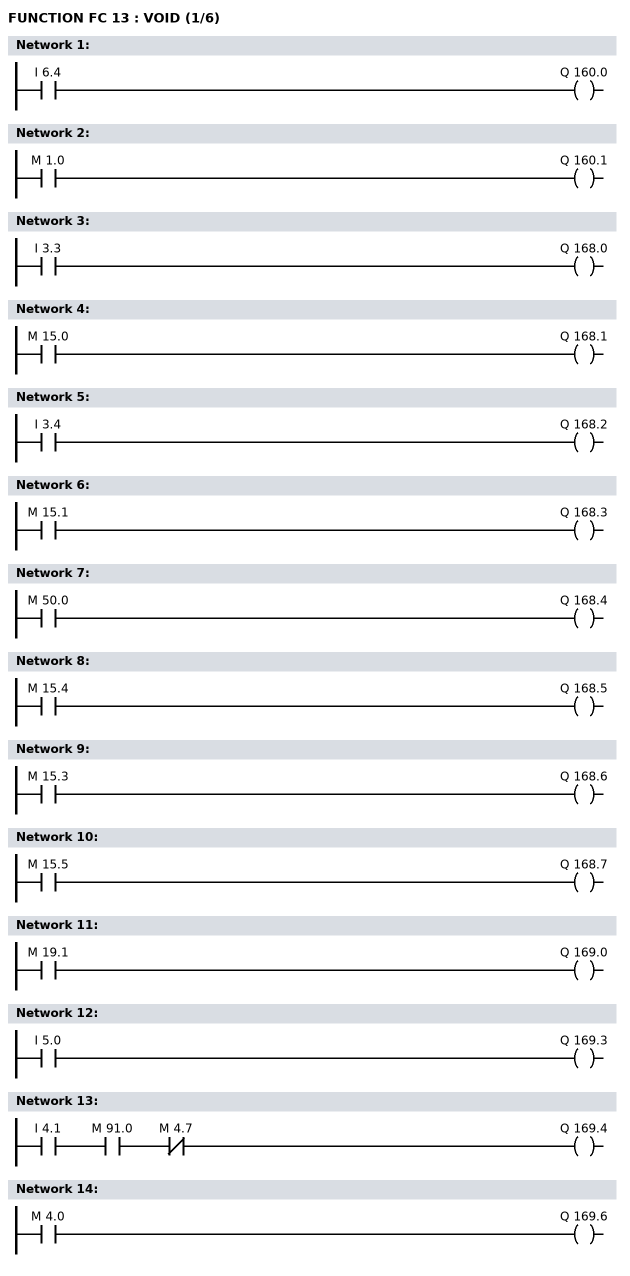

      A     I      6.4;
      =     Q    160.0;
NETWORK
TITLE =

      A     M      1.0;
      =     Q    160.1;
NETWORK
TITLE =

      A     I      3.3;
      =     Q    168.0;
NETWORK
TITLE =

      A     M     15.0;
      =     Q    168.1;
NETWORK
TITLE =

      A     I      3.4;
      =     Q    168.2;
NETWORK
TITLE =

      A     M     15.1;
      =     Q    168.3;
NETWORK
TITLE =

      A     M     50.0;
      =     Q    168.4;
NETWORK
TITLE =

      A     M     15.4;
      =     Q    168.5;
NETWORK
TITLE =

      A     M     15.3;
      =     Q    168.6;
NETWORK
TITLE =

      A     M     15.5;
      =     Q    168.7;
NETWORK
TITLE =

      A     M     19.1;
      =     Q    169.0;
NETWORK
TITLE =

      A     I      5.0;
      =     Q    169.3;
NETWORK
TITLE =

      A     I      4.1;
      A     M     91.0;
      AN    M      4.7;
      =     Q    169.4;
NETWORK
TITLE =

      A     M      4.0;
      =     Q    169.6;
NETWORK
TITLE =
